Staubli VAL3: utAppearance.dtx

public bool bVisibility
